(* IEC 61131-3 sources: 2026_Projet_YGO_ExcavatriceDragage/TOOLS/TEST_AUTO_CI/RESULTS/H_TREUILS_BENNE/tests (part 3) *)

(* ---- test_fb_winch.st ---- *)
(* =======================================================================
   🧪 test_fb_winch.st — FB_Winch (TC-P10-011, 017, 019, 042.1, 052.1, T216-AC4)
   ───────────────────────────────────────────────────────────────
   Fiche : DOC/AF/AF_Partie-10_Fonction_Winch/FB_Winch_v1.0.md
   Conventions : 1 appel fb() = 1 scan ; ADVANCE_TIME(10000000) entre les
   scans pour les fronts R_TRIG ; hex décrit en décimal (bit 0 = 1, bit 15 = 32768).
   Table valide : seuils croissants [10,30,50,70,90], P2..P5 au moins 1 contacteur TRUE.
   Interface structs : DriveRequest / Sensors / Config passés en variables
   (le harnais STruCpp ne supporte pas les littéraux de struct en appel FB).
   ======================================================================= *)

SETUP
VAR
    FB_W : FB_Winch;
    Table : ST_SpeedStepTable;
    DriveReq : ST_fbWinch_DriveRequest;
    Sens : ST_fbWinch_Sensors;
    Cfg : ST_fbWinch_Cfg;
END_VAR
END_SETUP

(* ── Table valide commune ── *)

TEST 'TC-P03-001 Dynamique Enable : neutralisation initiale, transition Ready au repos, puis coupure'
    Table.StepThreshold_Pct[1] := 10.0;
    Table.StepThreshold_Pct[2] := 30.0;
    Table.StepThreshold_Pct[3] := 50.0;
    Table.StepThreshold_Pct[4] := 70.0;
    Table.StepThreshold_Pct[5] := 90.0;
    Table.P2R1 := TRUE;
    Table.P3R1 := TRUE;
    Table.P4R1 := TRUE;
    Table.P5R1 := TRUE;
    Cfg.SpeedStepTable := Table;
    Sens.Homed := TRUE;
    Sens.ContactorsAllOff := TRUE;
    Sens.SpeedGuardReady := TRUE;

    (* Scan 0 : Enable=FALSE -> Neutralisation initiale *)
    DriveReq.RunRequest := FALSE;
    DriveReq.ReqAscent := FALSE; DriveReq.ReqDescend := FALSE;
    DriveReq.SpeedTgt_Pct := 0.0;
    FB_W(Enable := FALSE, Reset := FALSE, PowerContactorEngaged := TRUE,
         DriveRequest := DriveReq, Sensors := Sens, Config := Cfg);
    ASSERT_FALSE(FB_W.Ready, 'Enable=FALSE -> Ready=FALSE (neutralise)');

    ADVANCE_TIME(10000000);

    (* Scan 1 : Enable=TRUE -> Premier scan d initialisation *)
    FB_W(Enable := TRUE, Reset := FALSE, PowerContactorEngaged := TRUE,
         DriveRequest := DriveReq, Sensors := Sens, Config := Cfg);

    ADVANCE_TIME(10000000);

    (* Scan 2 : Regime nominal etabli -> Ready=TRUE *)
    FB_W(Enable := TRUE, Reset := FALSE, PowerContactorEngaged := TRUE,
         DriveRequest := DriveReq, Sensors := Sens, Config := Cfg);
    ASSERT_TRUE(FB_W.Ready, 'Enable=TRUE etabli -> Ready=TRUE (nominal)');

    ADVANCE_TIME(10000000);

    (* Scan 3 : Enable=FALSE -> Coupure nette et re-neutralisation *)
    FB_W(Enable := FALSE, Reset := FALSE, PowerContactorEngaged := TRUE,
         DriveRequest := DriveReq, Sensors := Sens, Config := Cfg);
    ASSERT_FALSE(FB_W.Ready, 'Enable=FALSE -> Ready retombe a FALSE');
END_TEST

TEST 'TC-P10-011 Inversion Fwd<->Rev : neutre->sens immediat, inversion exige delai + rampe a 0'
    Table.StepThreshold_Pct[1] := 10.0;
    Table.StepThreshold_Pct[2] := 30.0;
    Table.StepThreshold_Pct[3] := 50.0;
    Table.StepThreshold_Pct[4] := 70.0;
    Table.StepThreshold_Pct[5] := 90.0;
    Table.P2R1 := TRUE;
    Table.P3R1 := TRUE;
    Table.P4R1 := TRUE;
    Table.P5R1 := TRUE;
    Cfg.SpeedStepTable := Table;
    Sens.Homed := TRUE;
    Sens.ContactorsAllOff := TRUE;
    Sens.SpeedGuardReady := TRUE;

    (* Scan 1 : regime nominal *)
    DriveReq.RunRequest := FALSE;
    DriveReq.ReqAscent := FALSE; DriveReq.ReqDescend := FALSE;
    DriveReq.SpeedTgt_Pct := 0.0;
    FB_W(Enable := TRUE, Reset := FALSE, PowerContactorEngaged := TRUE,
         DriveRequest := DriveReq, Sensors := Sens, Config := Cfg);
    ADVANCE_TIME(10000000);
    FB_W(Enable := TRUE, Reset := FALSE, PowerContactorEngaged := TRUE,
         DriveRequest := DriveReq, Sensors := Sens, Config := Cfg);
    ASSERT_TRUE(FB_W.Ready, 'Treuil pret');

    (* Scan 2 : neutre -> montee = IMMEDIAT (pas de DirectionChangePending) *)
    ADVANCE_TIME(10000000);
    DriveReq.RunRequest := TRUE;
    DriveReq.ReqAscent := TRUE; DriveReq.ReqDescend := FALSE;
    DriveReq.SpeedTgt_Pct := 20.0;
    FB_W(Enable := TRUE, Reset := FALSE, PowerContactorEngaged := TRUE,
         DriveRequest := DriveReq, Sensors := Sens, Config := Cfg);
    ASSERT_EQ(FB_W.CommandedDirection, 1, 'Neutre->montee : CommandedDirection=1 immediat');
    ASSERT_FALSE(FB_W.DirectionChangePending, 'Neutre->montee : pas de pending');
    ASSERT_TRUE(FB_W.RelayFwd, 'Montee -> RelayFwd');

    (* Scan 3 : arret reel via neutre (StartStop=FALSE, Direction=0) -> StepNumber=0,
       CommandedDirection=0 (relais/diagnostic neutres) ; le dernier sens non nul est
       memorise en interne (LastDirection) pour l'interlock de reprise opposee *)
    ADVANCE_TIME(10000000);
    DriveReq.RunRequest := FALSE;
    DriveReq.ReqAscent := FALSE; DriveReq.ReqDescend := FALSE;
    DriveReq.SpeedTgt_Pct := 0.0;
    FB_W(Enable := TRUE, Reset := FALSE, PowerContactorEngaged := TRUE,
         DriveRequest := DriveReq, Sensors := Sens, Config := Cfg);
    ASSERT_EQ(FB_W.StepNumber, 0, 'Arret -> StepNumber=0');
    ASSERT_EQ(FB_W.CommandedDirection, 0, 'Arret via neutre : CommandedDirection=0 (relais/diagnostic neutres)');

    (* Scan 4 : inversion montee->descente apres neutre (StepNumber=0) -> pending + rampe a 0 *)
    ADVANCE_TIME(10000000);
    DriveReq.RunRequest := TRUE;
    DriveReq.ReqAscent := FALSE; DriveReq.ReqDescend := TRUE;
    DriveReq.SpeedTgt_Pct := 20.0;
    FB_W(Enable := TRUE, Reset := FALSE, PowerContactorEngaged := TRUE,
         DriveRequest := DriveReq, Sensors := Sens, Config := Cfg);
    ASSERT_TRUE(FB_W.DirectionChangePending, 'Inversion apres neutre -> DirectionChangePending=TRUE');
    ASSERT_EQ(FB_W.StepNumber, 0, 'Inversion : rampe forcee a 0 pendant attente');

    (* Scan 5 : apres DirectionInterlockDelayDescent=400ms -> CommandedDirection=-1 *)
    ADVANCE_TIME(400000000);
    FB_W(Enable := TRUE, Reset := FALSE, PowerContactorEngaged := TRUE,
         DriveRequest := DriveReq, Sensors := Sens, Config := Cfg);
    ASSERT_EQ(FB_W.CommandedDirection, -1, 'Apres 400ms -> CommandedDirection=-1');
    ASSERT_FALSE(FB_W.DirectionChangePending, 'Apres delai -> pending leve');
END_TEST

TEST 'TC-P10-011b Inversion via neutre : montee reelle -> relache neutre -> reprise descente -> temps mort + zero relais'
    Table.StepThreshold_Pct[1] := 10.0;
    Table.StepThreshold_Pct[2] := 30.0;
    Table.StepThreshold_Pct[3] := 50.0;
    Table.StepThreshold_Pct[4] := 70.0;
    Table.StepThreshold_Pct[5] := 90.0;
    Table.P2R1 := TRUE;
    Table.P3R1 := TRUE;
    Table.P4R1 := TRUE;
    Table.P5R1 := TRUE;
    Cfg.SpeedStepTable := Table;
    Sens.Homed := TRUE;
    Sens.ContactorsAllOff := TRUE;
    Sens.SpeedGuardReady := TRUE;

    (* Scan 1 : regime nominal *)
    DriveReq.RunRequest := FALSE;
    DriveReq.ReqAscent := FALSE; DriveReq.ReqDescend := FALSE;
    DriveReq.SpeedTgt_Pct := 0.0;
    FB_W(Enable := TRUE, Reset := FALSE, PowerContactorEngaged := TRUE,
         DriveRequest := DriveReq, Sensors := Sens, Config := Cfg);
    ADVANCE_TIME(10000000);
    FB_W(Enable := TRUE, Reset := FALSE, PowerContactorEngaged := TRUE,
         DriveRequest := DriveReq, Sensors := Sens, Config := Cfg);
    ASSERT_TRUE(FB_W.Ready, 'Treuil pret');

    (* Scan 2 : montee reelle etablie *)
    ADVANCE_TIME(10000000);
    DriveReq.RunRequest := TRUE;
    DriveReq.ReqAscent := TRUE; DriveReq.ReqDescend := FALSE;
    DriveReq.SpeedTgt_Pct := 90.0;
    FB_W(Enable := TRUE, Reset := FALSE, PowerContactorEngaged := TRUE,
         DriveRequest := DriveReq, Sensors := Sens, Config := Cfg);
    ASSERT_EQ(FB_W.CommandedDirection, 1, 'Montee reelle : CommandedDirection=1');
    ASSERT_TRUE(FB_W.RelayFwd, 'Montee reelle -> RelayFwd');

    (* Scan 3 : relachement neutre (Direction=0) -> StepNumber=0, CommandedDirection=0,
       relais coupes immediatement *)
    ADVANCE_TIME(10000000);
    DriveReq.RunRequest := FALSE;
    DriveReq.ReqAscent := FALSE; DriveReq.ReqDescend := FALSE;
    DriveReq.SpeedTgt_Pct := 0.0;
    FB_W(Enable := TRUE, Reset := FALSE, PowerContactorEngaged := TRUE,
         DriveRequest := DriveReq, Sensors := Sens, Config := Cfg);
    ASSERT_EQ(FB_W.StepNumber, 0, 'Neutre -> StepNumber=0');
    ASSERT_EQ(FB_W.CommandedDirection, 0, 'Neutre -> CommandedDirection=0 (relais/diagnostic neutres)');
    ASSERT_FALSE(FB_W.RelayFwd, 'Neutre -> RelayFwd coupe immediatement');
    ASSERT_FALSE(FB_W.RelayRev, 'Neutre -> RelayRev reste FALSE');

    (* Scan 4 : reprise descente (Direction=-1) -> pending + zero relais jusqu au delai *)
    ADVANCE_TIME(10000000);
    DriveReq.RunRequest := TRUE;
    DriveReq.ReqAscent := FALSE; DriveReq.ReqDescend := TRUE;
    DriveReq.SpeedTgt_Pct := 20.0;
    FB_W(Enable := TRUE, Reset := FALSE, PowerContactorEngaged := TRUE,
         DriveRequest := DriveReq, Sensors := Sens, Config := Cfg);
    ASSERT_TRUE(FB_W.DirectionChangePending, 'Reprise opposee apres neutre -> pending');
    ASSERT_EQ(FB_W.StepNumber, 0, 'Reprise opposee -> StepNumber=0 (rampe a 0)');
    ASSERT_FALSE(FB_W.RelayRev, 'Reprise opposee -> RelayRev retenu jusqu au delai');

    (* Scan 5 : apres DirectionInterlockDelayDescent=400ms -> CommandedDirection=-1, RelayRev *)
    ADVANCE_TIME(400000000);
    FB_W(Enable := TRUE, Reset := FALSE, PowerContactorEngaged := TRUE,
         DriveRequest := DriveReq, Sensors := Sens, Config := Cfg);
    ASSERT_EQ(FB_W.CommandedDirection, -1, 'Apres delai -> CommandedDirection=-1');
    ASSERT_FALSE(FB_W.DirectionChangePending, 'Apres delai -> pending leve');
    ASSERT_TRUE(FB_W.RelayRev, 'Apres delai -> RelayRev commande');
END_TEST

TEST 'TC-P10-011c Reprise du MEME sens apres neutre : depart immediat (pas de pending)'
    Table.StepThreshold_Pct[1] := 10.0;
    Table.StepThreshold_Pct[2] := 30.0;
    Table.StepThreshold_Pct[3] := 50.0;
    Table.StepThreshold_Pct[4] := 70.0;
    Table.StepThreshold_Pct[5] := 90.0;
    Table.P2R1 := TRUE;
    Table.P3R1 := TRUE;
    Table.P4R1 := TRUE;
    Table.P5R1 := TRUE;
    Cfg.SpeedStepTable := Table;
    Sens.Homed := TRUE;
    Sens.ContactorsAllOff := TRUE;
    Sens.SpeedGuardReady := TRUE;

    (* Scan 1 : regime nominal *)
    DriveReq.RunRequest := FALSE;
    DriveReq.ReqAscent := FALSE; DriveReq.ReqDescend := FALSE;
    DriveReq.SpeedTgt_Pct := 0.0;
    FB_W(Enable := TRUE, Reset := FALSE, PowerContactorEngaged := TRUE,
         DriveRequest := DriveReq, Sensors := Sens, Config := Cfg);
    ADVANCE_TIME(10000000);
    FB_W(Enable := TRUE, Reset := FALSE, PowerContactorEngaged := TRUE,
         DriveRequest := DriveReq, Sensors := Sens, Config := Cfg);
    ASSERT_TRUE(FB_W.Ready, 'Treuil pret');

    (* Scan 2 : montee reelle etablie *)
    ADVANCE_TIME(10000000);
    DriveReq.RunRequest := TRUE;
    DriveReq.ReqAscent := TRUE; DriveReq.ReqDescend := FALSE;
    DriveReq.SpeedTgt_Pct := 20.0;
    FB_W(Enable := TRUE, Reset := FALSE, PowerContactorEngaged := TRUE,
         DriveRequest := DriveReq, Sensors := Sens, Config := Cfg);
    ASSERT_EQ(FB_W.CommandedDirection, 1, 'Montee reelle : CommandedDirection=1');
    ASSERT_TRUE(FB_W.RelayFwd, 'Montee reelle -> RelayFwd');

    (* Scan 3 : relachement neutre -> CommandedDirection=0 *)
    ADVANCE_TIME(10000000);
    DriveReq.RunRequest := FALSE;
    DriveReq.ReqAscent := FALSE; DriveReq.ReqDescend := FALSE;
    DriveReq.SpeedTgt_Pct := 0.0;
    FB_W(Enable := TRUE, Reset := FALSE, PowerContactorEngaged := TRUE,
         DriveRequest := DriveReq, Sensors := Sens, Config := Cfg);
    ASSERT_EQ(FB_W.CommandedDirection, 0, 'Neutre -> CommandedDirection=0');

    (* Scan 4 : reprise du MEME sens (montee) -> depart immediat, pas de pending *)
    ADVANCE_TIME(10000000);
    DriveReq.RunRequest := TRUE;
    DriveReq.ReqAscent := TRUE; DriveReq.ReqDescend := FALSE;
    DriveReq.SpeedTgt_Pct := 20.0;
    FB_W(Enable := TRUE, Reset := FALSE, PowerContactorEngaged := TRUE,
         DriveRequest := DriveReq, Sensors := Sens, Config := Cfg);
    ASSERT_EQ(FB_W.CommandedDirection, 1, 'Reprise meme sens -> CommandedDirection=1 immediat');
    ASSERT_FALSE(FB_W.DirectionChangePending, 'Reprise meme sens -> pas de pending');
    ASSERT_TRUE(FB_W.RelayFwd, 'Reprise meme sens -> RelayFwd immediat');
END_TEST

TEST 'TC-P10-017 Config palier invalide : palier 0, sorties sures'
    (* Table invalide : seuils non croissants (tous a 0) *)
    Table.StepThreshold_Pct[1] := 0.0;
    Table.StepThreshold_Pct[2] := 0.0;
    Table.StepThreshold_Pct[3] := 0.0;
    Table.StepThreshold_Pct[4] := 0.0;
    Table.StepThreshold_Pct[5] := 0.0;
    Cfg.SpeedStepTable := Table;
    Sens.Homed := TRUE;
    Sens.ContactorsAllOff := TRUE;
    Sens.SpeedGuardReady := TRUE;

    (* Scan 1 : Enable=TRUE, config invalide -> ConfigError latche *)
    DriveReq.RunRequest := TRUE;
    DriveReq.ReqAscent := TRUE; DriveReq.ReqDescend := FALSE;
    DriveReq.SpeedTgt_Pct := 50.0;
    FB_W(Enable := TRUE, Reset := FALSE, PowerContactorEngaged := TRUE,
         DriveRequest := DriveReq, Sensors := Sens, Config := Cfg);
    ADVANCE_TIME(10000000);
    FB_W(Enable := TRUE, Reset := FALSE, PowerContactorEngaged := TRUE,
         DriveRequest := DriveReq, Sensors := Sens, Config := Cfg);
    ASSERT_TRUE(FB_W.Fault.Error, 'Config invalide -> Error');
    ASSERT_EQ(FB_W.StepNumber, 0, 'Config invalide -> palier 0');
    ASSERT_FALSE(FB_W.RelayFwd, 'Config invalide -> RelayFwd=FALSE (sortie sure)');
    ASSERT_FALSE(FB_W.RelayRev, 'Config invalide -> RelayRev=FALSE');
    ASSERT_FALSE(FB_W.Contactor1, 'Config invalide -> Contactor1=FALSE');
END_TEST

(* TC-P10-018 (StuckClosed) deplace/adapte dans test_fb_safety_winch.st (T181-02/03 AC5) :
   FB_Winch ne produit plus la detection contacteur colle — proprietaire unique FB_Safety_Winch. *)

TEST 'TC-P10-019 Ordre MainTask : Safety -> WinchControl -> PRG_06_Outputs'
    (* (essai site — stub) : l ordre d execution MainTask (Safety -> WinchControl -> PRG_06)
       est une propriete de la tache CODESYS, non automatisable en boite noire FB. On verifie
       ici la brique amont : FB_Winch produit bien sa demande sortie (RelayFwd) qui sera
       consommee par la barriere finale PRG_06. *)
    Table.StepThreshold_Pct[1] := 10.0;
    Table.StepThreshold_Pct[2] := 30.0;
    Table.StepThreshold_Pct[3] := 50.0;
    Table.StepThreshold_Pct[4] := 70.0;
    Table.StepThreshold_Pct[5] := 90.0;
    Table.P2R1 := TRUE;
    Table.P3R1 := TRUE;
    Table.P4R1 := TRUE;
    Table.P5R1 := TRUE;
    Cfg.SpeedStepTable := Table;
    Sens.Homed := TRUE;
    Sens.ContactorsAllOff := TRUE;
    Sens.SpeedGuardReady := TRUE;

    DriveReq.RunRequest := FALSE;
    DriveReq.ReqAscent := FALSE; DriveReq.ReqDescend := FALSE;
    DriveReq.SpeedTgt_Pct := 0.0;
    FB_W(Enable := TRUE, Reset := FALSE, PowerContactorEngaged := TRUE,
         DriveRequest := DriveReq, Sensors := Sens, Config := Cfg);
    ADVANCE_TIME(10000000);
    DriveReq.RunRequest := TRUE;
    DriveReq.ReqAscent := TRUE; DriveReq.ReqDescend := FALSE;
    DriveReq.SpeedTgt_Pct := 20.0;
    FB_W(Enable := TRUE, Reset := FALSE, PowerContactorEngaged := TRUE,
         DriveRequest := DriveReq, Sensors := Sens, Config := Cfg);
    ASSERT_TRUE(FB_W.RelayFwd, 'Demande montee produite (consommee par PRG_06)');
    ASSERT_TRUE(FB_W.Contactor1, 'Palier 1 demande');
END_TEST

TEST 'TC-P10-042.1 Plafonds dynamiques palier : descente max 3, montee max 5, approche capteur haut=1'
    Table.StepThreshold_Pct[1] := 10.0;
    Table.StepThreshold_Pct[2] := 30.0;
    Table.StepThreshold_Pct[3] := 50.0;
    Table.StepThreshold_Pct[4] := 70.0;
    Table.StepThreshold_Pct[5] := 90.0;
    Table.P2R1 := TRUE;
    Table.P3R1 := TRUE;
    Table.P4R1 := TRUE;
    Table.P5R1 := TRUE;
    Cfg.SpeedStepTable := Table;
    Sens.Homed := TRUE;
    Sens.ContactorsAllOff := TRUE;
    Sens.SpeedGuardReady := TRUE;
    DriveReq.HomingApproachActive := FALSE;
    Sens.CablePosM := 0.0;
    Cfg.SlowdownDistance_M := 1.0;

    (* Scan 1 : regime nominal *)
    DriveReq.RunRequest := FALSE;
    DriveReq.ReqAscent := FALSE; DriveReq.ReqDescend := FALSE;
    DriveReq.SpeedTgt_Pct := 0.0;
    FB_W(Enable := TRUE, Reset := FALSE, PowerContactorEngaged := TRUE,
         DriveRequest := DriveReq, Sensors := Sens, Config := Cfg);
    ADVANCE_TIME(10000000);
    FB_W(Enable := TRUE, Reset := FALSE, PowerContactorEngaged := TRUE,
         DriveRequest := DriveReq, Sensors := Sens, Config := Cfg);

    (* Descente : SpeedTgt_Pct=90 -> RequestedStep cape a CfgMaxStepDescente=3 *)
    ADVANCE_TIME(10000000);
    DriveReq.RunRequest := TRUE;
    DriveReq.ReqAscent := FALSE; DriveReq.ReqDescend := TRUE;
    DriveReq.SpeedTgt_Pct := 90.0;
    FB_W(Enable := TRUE, Reset := FALSE, PowerContactorEngaged := TRUE,
         DriveRequest := DriveReq, Sensors := Sens, Config := Cfg);
    ASSERT_EQ(FB_W.RequestedStep, 3, 'Descente : palier cape a 3 (CfgMaxStepDescente)');

    (* Reset + montee : SpeedTgt_Pct=90 -> RequestedStep=5 (MaxStepAscent) *)
    ADVANCE_TIME(10000000);
    DriveReq.RunRequest := FALSE;
    DriveReq.ReqAscent := FALSE; DriveReq.ReqDescend := FALSE;
    DriveReq.SpeedTgt_Pct := 0.0;
    FB_W(Enable := TRUE, Reset := TRUE, PowerContactorEngaged := TRUE,
         DriveRequest := DriveReq, Sensors := Sens, Config := Cfg);
    ADVANCE_TIME(10000000);
    DriveReq.RunRequest := TRUE;
    DriveReq.ReqAscent := TRUE; DriveReq.ReqDescend := FALSE;
    DriveReq.SpeedTgt_Pct := 90.0;
    FB_W(Enable := TRUE, Reset := FALSE, PowerContactorEngaged := TRUE,
         DriveRequest := DriveReq, Sensors := Sens, Config := Cfg);
    ASSERT_EQ(FB_W.RequestedStep, 5, 'Montee : palier 5 (MaxStepAscent)');

    (* Approche capteur haut : HomingApproachActive=TRUE -> palier 1 *)
    ADVANCE_TIME(10000000);
    DriveReq.RunRequest := FALSE;
    DriveReq.ReqAscent := FALSE; DriveReq.ReqDescend := FALSE;
    DriveReq.SpeedTgt_Pct := 0.0;
    FB_W(Enable := TRUE, Reset := TRUE, PowerContactorEngaged := TRUE,
         DriveRequest := DriveReq, Sensors := Sens, Config := Cfg);
    ADVANCE_TIME(10000000);
    DriveReq.RunRequest := TRUE;
    DriveReq.ReqAscent := TRUE; DriveReq.ReqDescend := FALSE;
    DriveReq.SpeedTgt_Pct := 90.0;
    DriveReq.HomingApproachActive := TRUE;
    FB_W(Enable := TRUE, Reset := FALSE, PowerContactorEngaged := TRUE,
         DriveRequest := DriveReq, Sensors := Sens, Config := Cfg);
    ASSERT_EQ(FB_W.RequestedStep, 1, 'Approche capteur haut : palier 1');

    (* Zone ralentissement haut : CablePosM >= TopLimitM - CfgSlowdownDistanceM -> palier 1 *)
    ADVANCE_TIME(10000000);
    DriveReq.RunRequest := FALSE;
    DriveReq.ReqAscent := FALSE; DriveReq.ReqDescend := FALSE;
    DriveReq.SpeedTgt_Pct := 0.0;
    DriveReq.HomingApproachActive := FALSE;
    FB_W(Enable := TRUE, Reset := TRUE, PowerContactorEngaged := TRUE,
         DriveRequest := DriveReq, Sensors := Sens, Config := Cfg);
    ADVANCE_TIME(10000000);
    DriveReq.RunRequest := TRUE;
    DriveReq.ReqAscent := TRUE; DriveReq.ReqDescend := FALSE;
    DriveReq.SpeedTgt_Pct := 90.0;
    DriveReq.TopLimitM := 8.5;
    Sens.CablePosM := 8.0;
    Cfg.SlowdownDistance_M := 1.0;
    FB_W(Enable := TRUE, Reset := FALSE, PowerContactorEngaged := TRUE,
         DriveRequest := DriveReq, Sensors := Sens, Config := Cfg);
    ASSERT_TRUE(FB_W.InTopSlowdownZone, 'Zone ralentissement haut active');
    ASSERT_EQ(FB_W.RequestedStep, 1, 'Zone ralentissement haut : palier 1');
END_TEST

TEST 'TC-P10-052.1 Garde-fou vitesse : vitesse non-stable -> palier 1 (activation par defaut)'
    (* (activation par defaut : T177) — SpeedGuardEnable est TRUE par defaut dans le code.
       On ne le force pas : le test verifie que le garde-fou est actif sans activation manuelle. *)
    Table.StepThreshold_Pct[1] := 10.0;
    Table.StepThreshold_Pct[2] := 30.0;
    Table.StepThreshold_Pct[3] := 50.0;
    Table.StepThreshold_Pct[4] := 70.0;
    Table.StepThreshold_Pct[5] := 90.0;
    Table.P2R1 := TRUE;
    Table.P3R1 := TRUE;
    Table.P4R1 := TRUE;
    Table.P5R1 := TRUE;
    Cfg.SpeedStepTable := Table;
    Sens.Homed := TRUE;
    Sens.ContactorsAllOff := TRUE;
    Sens.SpeedGuardReady := TRUE;
    DriveReq.HomingApproachActive := FALSE;
    Sens.CablePosM := 0.0;
    Cfg.SlowdownDistance_M := 1.0;

    (* Scan 1 : regime nominal *)
    DriveReq.RunRequest := FALSE;
    DriveReq.ReqAscent := FALSE; DriveReq.ReqDescend := FALSE;
    DriveReq.SpeedTgt_Pct := 0.0;
    FB_W(Enable := TRUE, Reset := FALSE, PowerContactorEngaged := TRUE,
         DriveRequest := DriveReq, Sensors := Sens, Config := Cfg);
    ADVANCE_TIME(10000000);
    FB_W(Enable := TRUE, Reset := FALSE, PowerContactorEngaged := TRUE,
         DriveRequest := DriveReq, Sensors := Sens, Config := Cfg);

    (* Scan 2 : SpeedGuardEnable=TRUE (defaut), SpeedGuardReady=FALSE (vitesse non stable) -> palier 1 *)
    ADVANCE_TIME(10000000);
    DriveReq.RunRequest := TRUE;
    DriveReq.ReqAscent := TRUE; DriveReq.ReqDescend := FALSE;
    DriveReq.SpeedTgt_Pct := 90.0;
    Sens.SpeedGuardReady := FALSE;
    FB_W(Enable := TRUE, Reset := FALSE, PowerContactorEngaged := TRUE,
         DriveRequest := DriveReq, Sensors := Sens, Config := Cfg);
    ASSERT_EQ(FB_W.RequestedStep, 1, 'Vitesse non stable -> palier 1 (garde-fou)');
    ASSERT_EQ(FB_W.StepNumber, 1, 'Vitesse non stable -> StepNumber=1');
END_TEST

(* ───────────────────────────────────────────────────────────────
   T216-AC4 : le plancher MinStepDown ne relance JAMAIS une descente
   lorsque le permis effectif de descente est FALSE (EffectiveSafeStop).
   REX : limite basse atteinte -> DescendPermit=FALSE -> la descente
   continuait au palier 1 (relance physique). Correction : gate du
   plancher par NOT EffectiveSafeStop (ligne 242 FB_Winch.st).
   ─────────────────────────────────────────────────────────────── *)

TEST 'T216-AC4-1 Regression : DescendPermit=FALSE + MinStepDown=1 -> StepNumber=0 et sorties=0'
    Table.StepThreshold_Pct[1] := 10.0;
    Table.StepThreshold_Pct[2] := 30.0;
    Table.StepThreshold_Pct[3] := 50.0;
    Table.StepThreshold_Pct[4] := 70.0;
    Table.StepThreshold_Pct[5] := 90.0;
    Table.P2R1 := TRUE;
    Table.P3R1 := TRUE;
    Table.P4R1 := TRUE;
    Table.P5R1 := TRUE;
    Cfg.SpeedStepTable := Table;
    Sens.Homed := TRUE;
    Sens.ContactorsAllOff := TRUE;
    Sens.SpeedGuardReady := TRUE;
    DriveReq.HomingApproachActive := FALSE;
    Sens.CablePosM := 0.0;
    Cfg.SlowdownDistance_M := 1.0;

    // Scan 1 : regime nominal neutre (arme l interlock direction), permis deja FALSE
    DriveReq.RunRequest := FALSE;
    DriveReq.ReqAscent := FALSE; DriveReq.ReqDescend := FALSE;
    DriveReq.SpeedStepReq := 0;
    DriveReq.MinStepDown := 1;
    DriveReq.MaxStepDown := 3;
    FB_W(Enable := TRUE, Reset := FALSE, PowerContactorEngaged := TRUE,
         DriveRequest := DriveReq, Sensors := Sens, Config := Cfg,
         SafeStop := FALSE, DescendPermit := FALSE, AscentPermit := TRUE);
    ADVANCE_TIME(10000000);
    FB_W(Enable := TRUE, Reset := FALSE, PowerContactorEngaged := TRUE,
         DriveRequest := DriveReq, Sensors := Sens, Config := Cfg,
         SafeStop := FALSE, DescendPermit := FALSE, AscentPermit := TRUE);

    // Scan 2 : operateur demande la descente (StartStop=TRUE, Dir=-1, SpeedStepReq=1)
    // MAIS DescendPermit=FALSE -> EffectiveSafeStop=TRUE doit garder RequestedStep=0.
    // Le plancher MinStepDown=1 ne doit PAS relever RequestedStep a >=1.
    ADVANCE_TIME(10000000);
    DriveReq.RunRequest := TRUE;
    DriveReq.ReqAscent := FALSE; DriveReq.ReqDescend := TRUE;
    DriveReq.SpeedStepReq := 1;
    FB_W(Enable := TRUE, Reset := FALSE, PowerContactorEngaged := TRUE,
         DriveRequest := DriveReq, Sensors := Sens, Config := Cfg,
         SafeStop := FALSE, DescendPermit := FALSE, AscentPermit := TRUE);
    ASSERT_EQ(FB_W.StepNumber, 0, 'Permis FALSE + MinStepDown : StepNumber=0 (descente interdite)');
    ASSERT_FALSE(FB_W.RelayFwd, 'Permis FALSE -> RelayFwd=FALSE');
    ASSERT_FALSE(FB_W.RelayRev, 'Permis FALSE -> RelayRev=FALSE (aucune relance descente)');
    ASSERT_FALSE(FB_W.Contactor1, 'Permis FALSE -> Contactor1=FALSE (sorties DQ descente = 0)');

    // Scan 3..4 : la demande est maintenue -> aucune relance palier apres cadence
    ADVANCE_TIME(10000000);
    FB_W(Enable := TRUE, Reset := FALSE, PowerContactorEngaged := TRUE,
         DriveRequest := DriveReq, Sensors := Sens, Config := Cfg,
         SafeStop := FALSE, DescendPermit := FALSE, AscentPermit := TRUE);
    ADVANCE_TIME(500000000);
    FB_W(Enable := TRUE, Reset := FALSE, PowerContactorEngaged := TRUE,
         DriveRequest := DriveReq, Sensors := Sens, Config := Cfg,
         SafeStop := FALSE, DescendPermit := FALSE, AscentPermit := TRUE);
    ASSERT_EQ(FB_W.StepNumber, 0, 'Permis FALSE : StepNumber reste 0 apres cadence (aucune relance)');
    ASSERT_FALSE(FB_W.RelayRev, 'Permis FALSE : RelayRev reste FALSE apres cadence');
END_TEST

TEST 'T216-AC4-2 Non-regression plongee Kobold : DescendPermit=TRUE + MinStepDown=3 -> plancher applique'
    Table.StepThreshold_Pct[1] := 10.0;
    Table.StepThreshold_Pct[2] := 30.0;
    Table.StepThreshold_Pct[3] := 50.0;
    Table.StepThreshold_Pct[4] := 70.0;
    Table.StepThreshold_Pct[5] := 90.0;
    Table.P2R1 := TRUE;
    Table.P3R1 := TRUE;
    Table.P4R1 := TRUE;
    Table.P5R1 := TRUE;
    Cfg.SpeedStepTable := Table;
    Sens.Homed := TRUE;
    Sens.ContactorsAllOff := TRUE;
    Sens.SpeedGuardReady := TRUE;
    DriveReq.HomingApproachActive := FALSE;
    Sens.CablePosM := 0.0;
    Cfg.SlowdownDistance_M := 1.0;

    // Scan 1 : regime nominal neutre
    DriveReq.RunRequest := FALSE;
    DriveReq.ReqAscent := FALSE; DriveReq.ReqDescend := FALSE;
    DriveReq.SpeedStepReq := 0;
    DriveReq.MinStepDown := 3;
    DriveReq.MaxStepDown := 3;
    FB_W(Enable := TRUE, Reset := FALSE, PowerContactorEngaged := TRUE,
         DriveRequest := DriveReq, Sensors := Sens, Config := Cfg,
         SafeStop := FALSE, DescendPermit := TRUE, AscentPermit := TRUE);
    ADVANCE_TIME(10000000);
    FB_W(Enable := TRUE, Reset := FALSE, PowerContactorEngaged := TRUE,
         DriveRequest := DriveReq, Sensors := Sens, Config := Cfg,
         SafeStop := FALSE, DescendPermit := TRUE, AscentPermit := TRUE);

    // Scan 2 : descente demandee, cible basse (SpeedStepReq=1) mais plancher MinStepDown=3
    // permis OK -> le plancher releve RequestedStep a 3 (clamp au plafond MaxStepDown=3)
    ADVANCE_TIME(10000000);
    DriveReq.RunRequest := TRUE;
    DriveReq.ReqAscent := FALSE; DriveReq.ReqDescend := TRUE;
    DriveReq.SpeedStepReq := 1;
    FB_W(Enable := TRUE, Reset := FALSE, PowerContactorEngaged := TRUE,
         DriveRequest := DriveReq, Sensors := Sens, Config := Cfg,
         SafeStop := FALSE, DescendPermit := TRUE, AscentPermit := TRUE);
    ASSERT_EQ(FB_W.RequestedStep, 3, 'Plancher MinStepDown=3 releve RequestedStep (permis OK)');
    ASSERT_TRUE(FB_W.StepNumber > 0, 'Plancher MinStepDown=3 -> StepNumber>0 (plongee maintenue)');
    ASSERT_TRUE(FB_W.RelayRev, 'Plancher MinStepDown=3 -> RelayRev commande (plongee Kobold)');

    // Scan 3..4 : cadence des 2 crans suivants (500ms/cran descente) -> StepNumber=3
    ADVANCE_TIME(500000000);
    FB_W(Enable := TRUE, Reset := FALSE, PowerContactorEngaged := TRUE,
         DriveRequest := DriveReq, Sensors := Sens, Config := Cfg,
         SafeStop := FALSE, DescendPermit := TRUE, AscentPermit := TRUE);
    ADVANCE_TIME(500000000);
    FB_W(Enable := TRUE, Reset := FALSE, PowerContactorEngaged := TRUE,
         DriveRequest := DriveReq, Sensors := Sens, Config := Cfg,
         SafeStop := FALSE, DescendPermit := TRUE, AscentPermit := TRUE);
    ASSERT_EQ(FB_W.StepNumber, 3, 'Cadence complet -> StepNumber=3 (plancher + plafond clamp)');
END_TEST

TEST 'T216-AC4-3 Perte du permis en mouvement : StepNumber retombe a 0 sans reprise de plancher'
    Table.StepThreshold_Pct[1] := 10.0;
    Table.StepThreshold_Pct[2] := 30.0;
    Table.StepThreshold_Pct[3] := 50.0;
    Table.StepThreshold_Pct[4] := 70.0;
    Table.StepThreshold_Pct[5] := 90.0;
    Table.P2R1 := TRUE;
    Table.P3R1 := TRUE;
    Table.P4R1 := TRUE;
    Table.P5R1 := TRUE;
    Cfg.SpeedStepTable := Table;
    Sens.Homed := TRUE;
    Sens.ContactorsAllOff := TRUE;
    Sens.SpeedGuardReady := TRUE;
    DriveReq.HomingApproachActive := FALSE;
    Sens.CablePosM := 0.0;
    Cfg.SlowdownDistance_M := 1.0;

    // Scan 1 : regime nominal neutre
    DriveReq.RunRequest := FALSE;
    DriveReq.ReqAscent := FALSE; DriveReq.ReqDescend := FALSE;
    DriveReq.SpeedStepReq := 0;
    DriveReq.MinStepDown := 1;
    DriveReq.MaxStepDown := 3;
    FB_W(Enable := TRUE, Reset := FALSE, PowerContactorEngaged := TRUE,
         DriveRequest := DriveReq, Sensors := Sens, Config := Cfg,
         SafeStop := FALSE, DescendPermit := TRUE, AscentPermit := TRUE);
    ADVANCE_TIME(10000000);
    FB_W(Enable := TRUE, Reset := FALSE, PowerContactorEngaged := TRUE,
         DriveRequest := DriveReq, Sensors := Sens, Config := Cfg,
         SafeStop := FALSE, DescendPermit := TRUE, AscentPermit := TRUE);

    // Scan 2-3 : descente etablie (permis OK) -> StepNumber=1, RelayRev commande
    ADVANCE_TIME(10000000);
    DriveReq.RunRequest := TRUE;
    DriveReq.ReqAscent := FALSE; DriveReq.ReqDescend := TRUE;
    DriveReq.SpeedStepReq := 1;
    FB_W(Enable := TRUE, Reset := FALSE, PowerContactorEngaged := TRUE,
         DriveRequest := DriveReq, Sensors := Sens, Config := Cfg,
         SafeStop := FALSE, DescendPermit := TRUE, AscentPermit := TRUE);
    ADVANCE_TIME(10000000);
    FB_W(Enable := TRUE, Reset := FALSE, PowerContactorEngaged := TRUE,
         DriveRequest := DriveReq, Sensors := Sens, Config := Cfg,
         SafeStop := FALSE, DescendPermit := TRUE, AscentPermit := TRUE);
    ASSERT_TRUE(FB_W.RelayRev, 'Pre-condition : descente etablie (permis OK)');

    // Scan 4..6 : le permis descente TOMBE (limite basse atteinte), l operateur maintient
    // la demande (StartStop=TRUE, Dir=-1, MinStepDown=1) -> StepNumber doit retomber a 0
    ADVANCE_TIME(10000000);
    FB_W(Enable := TRUE, Reset := FALSE, PowerContactorEngaged := TRUE,
         DriveRequest := DriveReq, Sensors := Sens, Config := Cfg,
         SafeStop := FALSE, DescendPermit := FALSE, AscentPermit := TRUE);
    ADVANCE_TIME(10000000);
    FB_W(Enable := TRUE, Reset := FALSE, PowerContactorEngaged := TRUE,
         DriveRequest := DriveReq, Sensors := Sens, Config := Cfg,
         SafeStop := FALSE, DescendPermit := FALSE, AscentPermit := TRUE);
    ADVANCE_TIME(10000000);
    FB_W(Enable := TRUE, Reset := FALSE, PowerContactorEngaged := TRUE,
         DriveRequest := DriveReq, Sensors := Sens, Config := Cfg,
         SafeStop := FALSE, DescendPermit := FALSE, AscentPermit := TRUE);
    ASSERT_EQ(FB_W.StepNumber, 0, 'Permis tombe en mouvement -> StepNumber retombe a 0');
    ASSERT_FALSE(FB_W.RelayRev, 'Permis tombe en mouvement -> RelayRev=FALSE (interruption descente)');

    // Scan 7-8 : maintien de la demande sans reprise -> aucune re-atterrissage palier
    ADVANCE_TIME(500000000);
    FB_W(Enable := TRUE, Reset := FALSE, PowerContactorEngaged := TRUE,
         DriveRequest := DriveReq, Sensors := Sens, Config := Cfg,
         SafeStop := FALSE, DescendPermit := FALSE, AscentPermit := TRUE);
    ADVANCE_TIME(500000000);
    FB_W(Enable := TRUE, Reset := FALSE, PowerContactorEngaged := TRUE,
         DriveRequest := DriveReq, Sensors := Sens, Config := Cfg,
         SafeStop := FALSE, DescendPermit := FALSE, AscentPermit := TRUE);
    ASSERT_EQ(FB_W.StepNumber, 0, 'Permis tombe : StepNumber reste 0 apres cadence (pas de reprise)');
    ASSERT_FALSE(FB_W.RelayRev, 'Permis tombe : RelayRev reste FALSE apres cadence');
END_TEST

(* ---- test_fb_winch_speed_learning.st ---- *)
(* =======================================================================
   🧪 test_fb_winch_speed_learning.st — FB_WinchSpeedLearning (T181-15)
   ───────────────────────────────────────────────────────────────
   Collecteur STRICTEMENT PASSIF des vitesses reelles par palier (RETAIN).
   Contrat : DOC/WFLOW/CONTRACTS/TASK_CONTRACT_T181-15_SPEED_LEARNING.yaml
   Conventions : 1 appel fb() = 1 scan ; Table est VAR_IN_OUT.
   ✅ Harnais copy-out (T181-21) : run_tests.py injecte le copy-out des
   VAR_IN_OUT apres chaque fb() (inject_var_in_out_copyout.py) — la variable
   de test Table reflete donc les ecritures du FB apres l'appel. On peut
   desormais asserter sur Table.Cell[...] (moyenne glissante + persistance
   RETAIN, TC-T181-15j).
   Strategie : pre-remplir la variable de test Table AVANT fb() pour les
   tests de frontiere/completude (a..i), et asserter sur Table.Cell[...]
   apres fb() pour prouver la moyenne glissante et la persistance RETAIN (j).
   Passivite (AC1/AC7) : verifiee par grep de l'interface FB (aucune sortie
   actionneur Relay* / Contactor* / Brake* / SpeedCmd ni Overspeed* / SpeedGuard* ).
   ======================================================================= *)

SETUP
VAR
    fb : FB_WinchSpeedLearning;
    Table : ST_fbWinchSpeedLearning_Table;
    Cfg : ST_fbWinchSpeedLearning_Cfg;
END_VAR
END_SETUP

(* ── Config commune : enveloppes par palier + MinSamples=3 ── *)

TEST 'TC-T181-15a LearnStart=FALSE : aucune collecte, table inchangee (AC3)'
    Cfg.MinSpeedMps[1] := 0.5; Cfg.MaxSpeedMps[1] := 2.0;
    Cfg.MinSpeedMps[2] := 1.0; Cfg.MaxSpeedMps[2] := 3.0;
    Cfg.MinSpeedMps[3] := 1.5; Cfg.MaxSpeedMps[3] := 4.0;
    Cfg.MinSpeedMps[4] := 2.0; Cfg.MaxSpeedMps[4] := 5.0;
    Cfg.MinSpeedMps[5] := 2.5; Cfg.MaxSpeedMps[5] := 6.0;
    Cfg.MinSamples := 3;

    (* Pre-remplissage : 1 cellule valide [1,1,1,1] *)
    Table.Cell[1][1][1][1].Valid := TRUE;
    Table.Cell[1][1][1][1].SpeedMps := 1.5;
    Table.Cell[1][1][1][1].SampleCount := 3;

    (* LearnStart=FALSE, toutes les autres conditions de collecte valides *)
    fb(Enable := TRUE, LearnStart := FALSE, WinchId := 1, Direction := 1,
       StepNumber := 1, MeasuredSpeedMps := 1.5, MeasuredSpeedValid := TRUE,
       LoadPresent := FALSE, StableForLearn := TRUE, Config := Cfg, Table := Table);

    ASSERT_FALSE(fb.Learning, 'LearnStart=FALSE : pas de collecte (Learning=FALSE)');
    ASSERT_FALSE(fb.LampLearn, 'LearnStart=FALSE : pas de voyant apprentissage');
    ASSERT_EQ(fb.CellsFilled, 1, 'LearnStart=FALSE : aucune nouvelle cellule (CellsFilled=1)');
END_TEST

TEST 'TC-T181-15b Conditions de collecte manquantes une a une : aucune ecriture (AC4)'
    Cfg.MinSpeedMps[1] := 0.5; Cfg.MaxSpeedMps[1] := 2.0;
    Cfg.MinSpeedMps[2] := 1.0; Cfg.MaxSpeedMps[2] := 3.0;
    Cfg.MinSpeedMps[3] := 1.5; Cfg.MaxSpeedMps[3] := 4.0;
    Cfg.MinSpeedMps[4] := 2.0; Cfg.MaxSpeedMps[4] := 5.0;
    Cfg.MinSpeedMps[5] := 2.5; Cfg.MaxSpeedMps[5] := 6.0;
    Cfg.MinSamples := 3;

    (* Mesure non valide : collecte bloquee -> aucune nouvelle cellule (CellsFilled reste 1) *)
    Table.Cell[1][1][1][1].Valid := TRUE;
    Table.Cell[1][1][1][1].SpeedMps := 1.5;
    Table.Cell[1][1][1][1].SampleCount := 3;
    fb(Enable := TRUE, LearnStart := TRUE, WinchId := 1, Direction := 1,
       StepNumber := 2, MeasuredSpeedMps := 1.5, MeasuredSpeedValid := FALSE,
       LoadPresent := FALSE, StableForLearn := TRUE, Config := Cfg, Table := Table);
    ASSERT_FALSE(fb.Learning, 'Mesure non valide : pas de collecte');
    ASSERT_EQ(fb.CellsFilled, 1, 'Mesure non valide : aucune nouvelle cellule');

    (* Conditions instables : collecte bloquee -> aucune nouvelle cellule *)
    Table.Cell[1][1][1][1].Valid := TRUE;
    Table.Cell[1][1][1][1].SpeedMps := 1.5;
    Table.Cell[1][1][1][1].SampleCount := 3;
    fb(Enable := TRUE, LearnStart := TRUE, WinchId := 1, Direction := 1,
       StepNumber := 3, MeasuredSpeedMps := 1.5, MeasuredSpeedValid := TRUE,
       LoadPresent := FALSE, StableForLearn := FALSE, Config := Cfg, Table := Table);
    ASSERT_FALSE(fb.Learning, 'Conditions instables : pas de collecte');
    ASSERT_EQ(fb.CellsFilled, 1, 'Conditions instables : aucune nouvelle cellule');

    (* Sens nul : collecte bloquee -> aucune nouvelle cellule *)
    Table.Cell[1][1][1][1].Valid := TRUE;
    Table.Cell[1][1][1][1].SpeedMps := 1.5;
    Table.Cell[1][1][1][1].SampleCount := 3;
    fb(Enable := TRUE, LearnStart := TRUE, WinchId := 1, Direction := 0,
       StepNumber := 4, MeasuredSpeedMps := 1.5, MeasuredSpeedValid := TRUE,
       LoadPresent := FALSE, StableForLearn := TRUE, Config := Cfg, Table := Table);
    ASSERT_FALSE(fb.Learning, 'Sens nul : pas de collecte');
    ASSERT_EQ(fb.CellsFilled, 1, 'Sens nul : aucune nouvelle cellule');

    (* Palier hors 1..5 : collecte bloquee -> aucune nouvelle cellule *)
    Table.Cell[1][1][1][1].Valid := TRUE;
    Table.Cell[1][1][1][1].SpeedMps := 1.5;
    Table.Cell[1][1][1][1].SampleCount := 3;
    fb(Enable := TRUE, LearnStart := TRUE, WinchId := 1, Direction := 1,
       StepNumber := 0, MeasuredSpeedMps := 1.5, MeasuredSpeedValid := TRUE,
       LoadPresent := FALSE, StableForLearn := TRUE, Config := Cfg, Table := Table);
    ASSERT_FALSE(fb.Learning, 'Palier hors 1..5 : pas de collecte');
    ASSERT_EQ(fb.CellsFilled, 1, 'Palier hors 1..5 : aucune nouvelle cellule');

    (* Axe hors 1..2 : collecte bloquee -> aucune nouvelle cellule *)
    Table.Cell[1][1][1][1].Valid := TRUE;
    Table.Cell[1][1][1][1].SpeedMps := 1.5;
    Table.Cell[1][1][1][1].SampleCount := 3;
    fb(Enable := TRUE, LearnStart := TRUE, WinchId := 0, Direction := 1,
       StepNumber := 1, MeasuredSpeedMps := 1.5, MeasuredSpeedValid := TRUE,
       LoadPresent := FALSE, StableForLearn := TRUE, Config := Cfg, Table := Table);
    ASSERT_FALSE(fb.Learning, 'Axe hors 1..2 : pas de collecte');
    ASSERT_EQ(fb.CellsFilled, 1, 'Axe hors 1..2 : aucune nouvelle cellule');
END_TEST

TEST 'TC-T181-15c Valid seulement a MinSamples : frontiere via CellsFilled (AC2/AC5)'
VAR
    i : INT;
    j : INT;
    k : INT;
    l : INT;
END_VAR
    Cfg.MinSpeedMps[1] := 0.5; Cfg.MaxSpeedMps[1] := 2.0;
    Cfg.MinSpeedMps[2] := 1.0; Cfg.MaxSpeedMps[2] := 3.0;
    Cfg.MinSpeedMps[3] := 1.5; Cfg.MaxSpeedMps[3] := 4.0;
    Cfg.MinSpeedMps[4] := 2.0; Cfg.MaxSpeedMps[4] := 5.0;
    Cfg.MinSpeedMps[5] := 2.5; Cfg.MaxSpeedMps[5] := 6.0;
    Cfg.MinSamples := 3;

    (* Part 1 : SampleCount=1 (MinSamples-2) -> apres 1 scan, encore < MinSamples -> non valide *)
    FOR i := 1 TO 2 DO
        FOR j := 1 TO 2 DO
            FOR k := 1 TO 2 DO
                FOR l := 1 TO 5 DO
                    Table.Cell[i][j][k][l].Valid := TRUE;
                END_FOR;
            END_FOR;
        END_FOR;
    END_FOR;
    Table.Cell[1][1][1][1].Valid := FALSE;
    Table.Cell[1][1][1][1].SampleCount := 1;
    Table.Cell[1][1][1][1].SpeedMps := 1.0;
    fb(Enable := TRUE, LearnStart := TRUE, WinchId := 1, Direction := 1,
       StepNumber := 1, MeasuredSpeedMps := 1.5, MeasuredSpeedValid := TRUE,
       LoadPresent := FALSE, StableForLearn := TRUE, Config := Cfg, Table := Table);
    ASSERT_EQ(fb.CellsFilled, 39, 'SampleCount 1->2 (<MinSamples) : cellule pas encore valide (39)');

    (* Part 2 : SampleCount=2 (MinSamples-1) -> apres 1 scan, MinSamples atteint -> valide *)
    FOR i := 1 TO 2 DO
        FOR j := 1 TO 2 DO
            FOR k := 1 TO 2 DO
                FOR l := 1 TO 5 DO
                    Table.Cell[i][j][k][l].Valid := TRUE;
                END_FOR;
            END_FOR;
        END_FOR;
    END_FOR;
    Table.Cell[1][1][1][1].Valid := FALSE;
    Table.Cell[1][1][1][1].SampleCount := 2;
    Table.Cell[1][1][1][1].SpeedMps := 1.0;
    fb(Enable := TRUE, LearnStart := TRUE, WinchId := 1, Direction := 1,
       StepNumber := 1, MeasuredSpeedMps := 1.5, MeasuredSpeedValid := TRUE,
       LoadPresent := FALSE, StableForLearn := TRUE, Config := Cfg, Table := Table);
    ASSERT_EQ(fb.CellsFilled, 40, 'SampleCount 2->3 (=MinSamples) : cellule validee (40)');
    ASSERT_TRUE(fb.TableComplete, 'MinSamples atteint sur la derniere cellule : TableComplete=TRUE');
END_TEST

TEST 'TC-T181-15d Hors enveloppe : cellule invalidee (Valid=FALSE, SampleCount=0, SpeedMps=0) (AC5)'
    Cfg.MinSpeedMps[1] := 0.5; Cfg.MaxSpeedMps[1] := 2.0;
    Cfg.MinSpeedMps[2] := 1.0; Cfg.MaxSpeedMps[2] := 3.0;
    Cfg.MinSpeedMps[3] := 1.5; Cfg.MaxSpeedMps[3] := 4.0;
    Cfg.MinSpeedMps[4] := 2.0; Cfg.MaxSpeedMps[4] := 5.0;
    Cfg.MinSpeedMps[5] := 2.5; Cfg.MaxSpeedMps[5] := 6.0;
    Cfg.MinSamples := 3;

    (* Cellule validee [1,1,1,1] puis injection hors enveloppe haute (5.0 > Max[1]=2.0) *)
    Table.Cell[1][1][1][1].Valid := TRUE;
    Table.Cell[1][1][1][1].SpeedMps := 1.5;
    Table.Cell[1][1][1][1].SampleCount := 3;
    fb(Enable := TRUE, LearnStart := TRUE, WinchId := 1, Direction := 1,
       StepNumber := 1, MeasuredSpeedMps := 5.0, MeasuredSpeedValid := TRUE,
       LoadPresent := FALSE, StableForLearn := TRUE, Config := Cfg, Table := Table);
    ASSERT_EQ(fb.CellsFilled, 0, 'Hors enveloppe haute : cellule invalidee (CellsFilled=0)');

    (* Injection sous la borne basse (0.4 < Min[1]=0.5) -> invalidation aussi *)
    Table.Cell[1][1][1][1].Valid := TRUE;
    Table.Cell[1][1][1][1].SpeedMps := 1.5;
    Table.Cell[1][1][1][1].SampleCount := 3;
    fb(Enable := TRUE, LearnStart := TRUE, WinchId := 1, Direction := 1,
       StepNumber := 1, MeasuredSpeedMps := 0.4, MeasuredSpeedValid := TRUE,
       LoadPresent := FALSE, StableForLearn := TRUE, Config := Cfg, Table := Table);
    ASSERT_EQ(fb.CellsFilled, 0, 'Sous borne basse : cellule invalidee (CellsFilled=0)');

    (* Borne exacte ==Max (2.0, inclusive) -> cellule conservee validee *)
    Table.Cell[1][1][1][1].Valid := TRUE;
    Table.Cell[1][1][1][1].SpeedMps := 1.5;
    Table.Cell[1][1][1][1].SampleCount := 3;
    fb(Enable := TRUE, LearnStart := TRUE, WinchId := 1, Direction := 1,
       StepNumber := 1, MeasuredSpeedMps := 2.0, MeasuredSpeedValid := TRUE,
       LoadPresent := FALSE, StableForLearn := TRUE, Config := Cfg, Table := Table);
    ASSERT_EQ(fb.CellsFilled, 1, 'Borne ==Max (2.0) inclusive : cellule conservee validee (1)');

    (* Borne exacte ==Min (0.5, inclusive) -> cellule conservee validee *)
    Table.Cell[1][1][1][1].Valid := TRUE;
    Table.Cell[1][1][1][1].SpeedMps := 1.5;
    Table.Cell[1][1][1][1].SampleCount := 3;
    fb(Enable := TRUE, LearnStart := TRUE, WinchId := 1, Direction := 1,
       StepNumber := 1, MeasuredSpeedMps := 0.5, MeasuredSpeedValid := TRUE,
       LoadPresent := FALSE, StableForLearn := TRUE, Config := Cfg, Table := Table);
    ASSERT_EQ(fb.CellsFilled, 1, 'Borne ==Min (0.5) inclusive : cellule conservee validee (1)');
END_TEST

TEST 'TC-T181-15e TableComplete : FALSE si une cellule manque, TRUE avec 40 cellules valides (AC6)'
VAR
    i : INT;
    j : INT;
    k : INT;
    l : INT;
END_VAR
    Cfg.MinSpeedMps[1] := 0.5; Cfg.MaxSpeedMps[1] := 2.0;
    Cfg.MinSpeedMps[2] := 1.0; Cfg.MaxSpeedMps[2] := 3.0;
    Cfg.MinSpeedMps[3] := 1.5; Cfg.MaxSpeedMps[3] := 4.0;
    Cfg.MinSpeedMps[4] := 2.0; Cfg.MaxSpeedMps[4] := 5.0;
    Cfg.MinSpeedMps[5] := 2.5; Cfg.MaxSpeedMps[5] := 6.0;
    Cfg.MinSamples := 1;

    (* Table partielle : 39 cellules valides, [2,2,2,5] manquante -> FALSE *)
    FOR i := 1 TO 2 DO
        FOR j := 1 TO 2 DO
            FOR k := 1 TO 2 DO
                FOR l := 1 TO 5 DO
                    Table.Cell[i][j][k][l].Valid := TRUE;
                END_FOR;
            END_FOR;
        END_FOR;
    END_FOR;
    Table.Cell[2][2][2][5].Valid := FALSE;

    fb(Enable := TRUE, LearnStart := FALSE, WinchId := 1, Direction := 1,
       StepNumber := 1, MeasuredSpeedMps := 1.0, MeasuredSpeedValid := TRUE,
       LoadPresent := FALSE, StableForLearn := TRUE, Config := Cfg, Table := Table);
    ASSERT_FALSE(fb.TableComplete, 'Table partielle (39/40) : TableComplete=FALSE');
    ASSERT_EQ(fb.CellsFilled, 39, 'Table partielle : CellsFilled=39');
    ASSERT_EQ(fb.CellsTotal, 40, 'CellsTotal=40 (2x2x2x5)');

    (* Table complete : 40 cellules valides -> TRUE *)
    Table.Cell[2][2][2][5].Valid := TRUE;
    fb(Enable := TRUE, LearnStart := FALSE, WinchId := 1, Direction := 1,
       StepNumber := 1, MeasuredSpeedMps := 1.0, MeasuredSpeedValid := TRUE,
       LoadPresent := FALSE, StableForLearn := TRUE, Config := Cfg, Table := Table);
    ASSERT_TRUE(fb.TableComplete, 'Table complete (40/40) : TableComplete=TRUE');
    ASSERT_EQ(fb.CellsFilled, 40, 'Table complete : CellsFilled=40');
END_TEST

TEST 'TC-T181-15f Passivite : sorties limitees au statut/diagnostic, aucune commande moteur (AC1/AC7)'
    (* La passivite (aucune sortie actionneur Relay* / Contactor* / Brake* / SpeedCmd ni
       Overspeed* / SpeedGuard* ) est verifiee par grep de l interface FB (AC1/AC7).
       Ce test confirme le comportement observable : pendant la collecte, seules les
       sorties de statut/diagnostic evoluent (Ready/Learning/LampLearn) + la Table. *)
    Cfg.MinSpeedMps[1] := 0.5; Cfg.MaxSpeedMps[1] := 2.0;
    Cfg.MinSpeedMps[2] := 1.0; Cfg.MaxSpeedMps[2] := 3.0;
    Cfg.MinSpeedMps[3] := 1.5; Cfg.MaxSpeedMps[3] := 4.0;
    Cfg.MinSpeedMps[4] := 2.0; Cfg.MaxSpeedMps[4] := 5.0;
    Cfg.MinSpeedMps[5] := 2.5; Cfg.MaxSpeedMps[5] := 6.0;
    Cfg.MinSamples := 3;

    fb(Enable := TRUE, LearnStart := TRUE, WinchId := 1, Direction := 1,
       StepNumber := 1, MeasuredSpeedMps := 1.0, MeasuredSpeedValid := TRUE,
       LoadPresent := FALSE, StableForLearn := TRUE, Config := Cfg, Table := Table);
    ASSERT_TRUE(fb.Ready, 'Enable=TRUE -> Ready=TRUE');
    ASSERT_TRUE(fb.Learning, 'Collecte active -> Learning=TRUE');
    ASSERT_TRUE(fb.LampLearn, 'Collecte active -> LampLearn=TRUE');
    ASSERT_EQ(fb.CellsTotal, 40, 'CellsTotal=40 (diagnostic)');

    (* Relache : Enable=FALSE -> Ready=FALSE, plus de collecte *)
    fb(Enable := FALSE, LearnStart := TRUE, WinchId := 1, Direction := 1,
       StepNumber := 1, MeasuredSpeedMps := 1.0, MeasuredSpeedValid := TRUE,
       LoadPresent := FALSE, StableForLearn := TRUE, Config := Cfg, Table := Table);
    ASSERT_FALSE(fb.Ready, 'Enable=FALSE -> Ready=FALSE');
    ASSERT_FALSE(fb.Learning, 'Enable=FALSE -> Learning=FALSE');
END_TEST

TEST 'TC-T181-15g Sens descente : cellule descente [1,2,1,1] ecrite, montee inchangee (AC2)'
VAR
    i : INT;
    j : INT;
    k : INT;
    l : INT;
END_VAR
    Cfg.MinSpeedMps[1] := 0.5; Cfg.MaxSpeedMps[1] := 2.0;
    Cfg.MinSpeedMps[2] := 1.0; Cfg.MaxSpeedMps[2] := 3.0;
    Cfg.MinSpeedMps[3] := 1.5; Cfg.MaxSpeedMps[3] := 4.0;
    Cfg.MinSpeedMps[4] := 2.0; Cfg.MaxSpeedMps[4] := 5.0;
    Cfg.MinSpeedMps[5] := 2.5; Cfg.MaxSpeedMps[5] := 6.0;
    Cfg.MinSamples := 1;

    (* 39 cellules valides, descente [1,2,1,1] vide. Direction=-1 -> SensIdx=2 *)
    FOR i := 1 TO 2 DO
        FOR j := 1 TO 2 DO
            FOR k := 1 TO 2 DO
                FOR l := 1 TO 5 DO
                    Table.Cell[i][j][k][l].Valid := TRUE;
                END_FOR;
            END_FOR;
        END_FOR;
    END_FOR;
    Table.Cell[1][2][1][1].Valid := FALSE;

    fb(Enable := TRUE, LearnStart := TRUE, WinchId := 1, Direction := -1,
       StepNumber := 1, MeasuredSpeedMps := 1.0, MeasuredSpeedValid := TRUE,
       LoadPresent := FALSE, StableForLearn := TRUE, Config := Cfg, Table := Table);
    ASSERT_EQ(fb.CellsFilled, 40, 'Descente : cellule descente [1,2,1,1] ecrite et validee (40)');
    ASSERT_TRUE(fb.TableComplete, 'Descente : table complete apres ecriture descente');
END_TEST

TEST 'TC-T181-15h Charge presente : cellule charge [1,1,2,1] ecrite, vide inchangee (AC2)'
VAR
    i : INT;
    j : INT;
    k : INT;
    l : INT;
END_VAR
    Cfg.MinSpeedMps[1] := 0.5; Cfg.MaxSpeedMps[1] := 2.0;
    Cfg.MinSpeedMps[2] := 1.0; Cfg.MaxSpeedMps[2] := 3.0;
    Cfg.MinSpeedMps[3] := 1.5; Cfg.MaxSpeedMps[3] := 4.0;
    Cfg.MinSpeedMps[4] := 2.0; Cfg.MaxSpeedMps[4] := 5.0;
    Cfg.MinSpeedMps[5] := 2.5; Cfg.MaxSpeedMps[5] := 6.0;
    Cfg.MinSamples := 1;

    (* 39 cellules valides, charge [1,1,2,1] vide. LoadPresent=TRUE -> ChargeIdx=2 *)
    FOR i := 1 TO 2 DO
        FOR j := 1 TO 2 DO
            FOR k := 1 TO 2 DO
                FOR l := 1 TO 5 DO
                    Table.Cell[i][j][k][l].Valid := TRUE;
                END_FOR;
            END_FOR;
        END_FOR;
    END_FOR;
    Table.Cell[1][1][2][1].Valid := FALSE;

    fb(Enable := TRUE, LearnStart := TRUE, WinchId := 1, Direction := 1,
       StepNumber := 1, MeasuredSpeedMps := 1.0, MeasuredSpeedValid := TRUE,
       LoadPresent := TRUE, StableForLearn := TRUE, Config := Cfg, Table := Table);
    ASSERT_EQ(fb.CellsFilled, 40, 'Charge : cellule charge [1,1,2,1] ecrite et validee (40)');
    ASSERT_TRUE(fb.TableComplete, 'Charge : table complete apres ecriture charge');
END_TEST

TEST 'TC-T181-15i Axe M2 (WinchId=2) : cellule [2,1,1,1] ecrite, M1 inchangee (AC2)'
VAR
    i : INT;
    j : INT;
    k : INT;
    l : INT;
END_VAR
    Cfg.MinSpeedMps[1] := 0.5; Cfg.MaxSpeedMps[1] := 2.0;
    Cfg.MinSpeedMps[2] := 1.0; Cfg.MaxSpeedMps[2] := 3.0;
    Cfg.MinSpeedMps[3] := 1.5; Cfg.MaxSpeedMps[3] := 4.0;
    Cfg.MinSpeedMps[4] := 2.0; Cfg.MaxSpeedMps[4] := 5.0;
    Cfg.MinSpeedMps[5] := 2.5; Cfg.MaxSpeedMps[5] := 6.0;
    Cfg.MinSamples := 1;

    (* 39 cellules valides, M2 [2,1,1,1] vide. WinchId=2 -> AxeIdx=2 *)
    FOR i := 1 TO 2 DO
        FOR j := 1 TO 2 DO
            FOR k := 1 TO 2 DO
                FOR l := 1 TO 5 DO
                    Table.Cell[i][j][k][l].Valid := TRUE;
                END_FOR;
            END_FOR;
        END_FOR;
    END_FOR;
    Table.Cell[2][1][1][1].Valid := FALSE;

    fb(Enable := TRUE, LearnStart := TRUE, WinchId := 2, Direction := 1,
       StepNumber := 1, MeasuredSpeedMps := 1.0, MeasuredSpeedValid := TRUE,
       LoadPresent := FALSE, StableForLearn := TRUE, Config := Cfg, Table := Table);
    ASSERT_EQ(fb.CellsFilled, 40, 'M2 : cellule [2,1,1,1] ecrite et validee (40)');
    ASSERT_TRUE(fb.TableComplete, 'M2 : table complete apres ecriture M2');
END_TEST

TEST 'TC-T181-15j Moyenne glissante + persistance RETAIN via copy-out (AC2)'
    (* Copy-out (T181-21) : apres fb(), la variable de test Table reflete les
       ecritures du FB sur la VAR_IN_OUT. On prouve ici la moyenne glissante
       (SpeedMps) et la persistance RETAIN (accumulation d'un scan a l'autre). *)
    Cfg.MinSpeedMps[1] := 0.5; Cfg.MaxSpeedMps[1] := 2.0;
    Cfg.MinSpeedMps[2] := 1.0; Cfg.MaxSpeedMps[2] := 3.0;
    Cfg.MinSpeedMps[3] := 1.5; Cfg.MaxSpeedMps[3] := 4.0;
    Cfg.MinSpeedMps[4] := 2.0; Cfg.MaxSpeedMps[4] := 5.0;
    Cfg.MinSpeedMps[5] := 2.5; Cfg.MaxSpeedMps[5] := 6.0;
    Cfg.MinSamples := 3;

    (* Cellule [1,1,1,1] vide. 1er echantillon 1.0 (plausible) -> SpeedMps=1.0, SampleCount=1 *)
    fb(Enable := TRUE, LearnStart := TRUE, WinchId := 1, Direction := 1,
       StepNumber := 1, MeasuredSpeedMps := 1.0, MeasuredSpeedValid := TRUE,
       LoadPresent := FALSE, StableForLearn := TRUE, Config := Cfg, Table := Table);
    ASSERT_EQ(Table.Cell[1][1][1][1].SampleCount, 1, '1er scan : SampleCount=1');
    ASSERT_NEAR(Table.Cell[1][1][1][1].SpeedMps, 1.0, 0.0001, '1er scan : SpeedMps=1.0');
    ASSERT_FALSE(Table.Cell[1][1][1][1].Valid, '1er scan : SampleCount<MinSamples -> Valid=FALSE');

    (* 2e echantillon 1.5 -> moyenne (1.0+1.5)/2 = 1.25, SampleCount=2 *)
    fb(Enable := TRUE, LearnStart := TRUE, WinchId := 1, Direction := 1,
       StepNumber := 1, MeasuredSpeedMps := 1.5, MeasuredSpeedValid := TRUE,
       LoadPresent := FALSE, StableForLearn := TRUE, Config := Cfg, Table := Table);
    ASSERT_EQ(Table.Cell[1][1][1][1].SampleCount, 2, '2e scan : SampleCount=2');
    ASSERT_NEAR(Table.Cell[1][1][1][1].SpeedMps, 1.25, 0.0001, '2e scan : moyenne (1.0+1.5)/2=1.25');
    ASSERT_FALSE(Table.Cell[1][1][1][1].Valid, '2e scan : SampleCount<MinSamples -> Valid=FALSE');

    (* 3e echantillon 1.5 -> moyenne (1.25*2+1.5)/3 = 1.3333, SampleCount=3 -> Valid *)
    fb(Enable := TRUE, LearnStart := TRUE, WinchId := 1, Direction := 1,
       StepNumber := 1, MeasuredSpeedMps := 1.5, MeasuredSpeedValid := TRUE,
       LoadPresent := FALSE, StableForLearn := TRUE, Config := Cfg, Table := Table);
    ASSERT_EQ(Table.Cell[1][1][1][1].SampleCount, 3, '3e scan : SampleCount=3');
    ASSERT_NEAR(Table.Cell[1][1][1][1].SpeedMps, 1.3333, 0.0001, '3e scan : moyenne (1.25*2+1.5)/3=1.3333');
    ASSERT_TRUE(Table.Cell[1][1][1][1].Valid, '3e scan : MinSamples atteint -> Valid=TRUE');
END_TEST

(* ---- test_fb_winch_symmetry.st ---- *)
(* =======================================================================
   test_fb_winch_symmetry.st -- T181-18 D11 : macro TC FB_Winch_Symmetry (F10.06)
   Observateur passif de symetrie / synchronisme M1-M2. Aucune action securite.
   Qualification : commande stable des 2 treuils, meme sens, au-dela de
   MinimumCommandTime_Ms (defaut 1000 ms) et vitesse au-dessus de MinimumSpeed_Mps.
   Les ecarts sont calcules a l arret.
   ======================================================================= *)

SETUP
VAR
    fb  : FB_Winch_Symmetry;
    Cfg : ST_fbWinch_Symmetry_Cfg;
    Dat : ST_fbWinch_Symmetry_Data;
END_VAR
END_SETUP

TEST 'TC-P10-T181-18a Cycle symetrique -> SymmetryValid et SymmetryOk'
    Cfg.MinimumCommandTime_Ms := 300;
    Cfg.MinimumSpeed_Mps := 0.05;
    Cfg.DeltaStartDelay_Ms := 100; Cfg.DeltaBrakeReleaseTime_Ms := 100;
    Cfg.DeltaBrakeApplyTime_Ms := 100; Cfg.DeltaStopDistance_Mm := 100;
    Cfg.DeltaStopTime_Ms := 200;
    fb(Reset := TRUE, M1CommandActive := FALSE, M2CommandActive := FALSE, M1Direction := 0, M2Direction := 0,
       M1BrakeCmd := FALSE, M2BrakeCmd := FALSE, M1BrakeApplied := TRUE, M2BrakeApplied := TRUE,
       M1Position_M := 0.0, M2Position_M := 0.0, M1Speed_Mps := 0.0, M2Speed_Mps := 0.0,
       SyncDeviation_M := 0.0, Config := Cfg, Data := Dat);
    fb(Reset := FALSE, M1CommandActive := TRUE, M2CommandActive := TRUE, M1Direction := 1, M2Direction := 1,
       M1BrakeCmd := TRUE, M2BrakeCmd := TRUE, M1BrakeApplied := FALSE, M2BrakeApplied := FALSE,
       M1Position_M := 0.0, M2Position_M := 0.0, M1Speed_Mps := 1.0, M2Speed_Mps := 1.0,
       SyncDeviation_M := 0.10, Config := Cfg, Data := Dat);
    ADVANCE_TIME(500000000);
    fb(Reset := FALSE, M1CommandActive := TRUE, M2CommandActive := TRUE, M1Direction := 1, M2Direction := 1,
       M1BrakeCmd := TRUE, M2BrakeCmd := TRUE, M1BrakeApplied := FALSE, M2BrakeApplied := FALSE,
       M1Position_M := 0.5, M2Position_M := 0.5, M1Speed_Mps := 1.0, M2Speed_Mps := 1.0,
       SyncDeviation_M := 0.10, Config := Cfg, Data := Dat);
    ADVANCE_TIME(500000000);
    fb(Reset := FALSE, M1CommandActive := TRUE, M2CommandActive := TRUE, M1Direction := 1, M2Direction := 1,
       M1BrakeCmd := TRUE, M2BrakeCmd := TRUE, M1BrakeApplied := FALSE, M2BrakeApplied := FALSE,
       M1Position_M := 1.0, M2Position_M := 1.0, M1Speed_Mps := 1.0, M2Speed_Mps := 1.0,
       SyncDeviation_M := 0.10, Config := Cfg, Data := Dat);
    ADVANCE_TIME(500000000);
    fb(Reset := FALSE, M1CommandActive := TRUE, M2CommandActive := TRUE, M1Direction := 1, M2Direction := 1,
       M1BrakeCmd := TRUE, M2BrakeCmd := TRUE, M1BrakeApplied := FALSE, M2BrakeApplied := FALSE,
       M1Position_M := 1.5, M2Position_M := 1.5, M1Speed_Mps := 1.0, M2Speed_Mps := 1.0,
       SyncDeviation_M := 0.10, Config := Cfg, Data := Dat);
    ADVANCE_TIME(500000000);
    fb(Reset := FALSE, M1CommandActive := FALSE, M2CommandActive := FALSE, M1Direction := 1, M2Direction := 1,
       M1BrakeCmd := FALSE, M2BrakeCmd := FALSE, M1BrakeApplied := TRUE, M2BrakeApplied := TRUE,
       M1Position_M := 2.0, M2Position_M := 2.0, M1Speed_Mps := 0.0, M2Speed_Mps := 0.0,
       SyncDeviation_M := 0.0, Config := Cfg, Data := Dat);
    ADVANCE_TIME(10000000);
    fb(Reset := FALSE, M1CommandActive := FALSE, M2CommandActive := FALSE, M1Direction := 1, M2Direction := 1,
       M1BrakeCmd := FALSE, M2BrakeCmd := FALSE, M1BrakeApplied := TRUE, M2BrakeApplied := TRUE,
       M1Position_M := 2.0, M2Position_M := 2.0, M1Speed_Mps := 0.0, M2Speed_Mps := 0.0,
       SyncDeviation_M := 0.0, Config := Cfg, Data := Dat);
    ASSERT_TRUE(fb.SymmetryValid, 'Cycle complet qualifie puis arrete -> mesure valide');
    ASSERT_TRUE(fb.SymmetryOk, 'M1 et M2 identiques -> tous les ecarts sous les seuils');
END_TEST

TEST 'TC-P10-T181-18b Reset remet les mesures a zero'
    Cfg.MinimumCommandTime_Ms := 300;
    Cfg.MinimumSpeed_Mps := 0.05;
    Cfg.DeltaStartDelay_Ms := 100; Cfg.DeltaBrakeReleaseTime_Ms := 100;
    Cfg.DeltaBrakeApplyTime_Ms := 100; Cfg.DeltaStopDistance_Mm := 100;
    Cfg.DeltaStopTime_Ms := 200;
    fb(Reset := TRUE, M1CommandActive := FALSE, M2CommandActive := FALSE, M1Direction := 0, M2Direction := 0,
       M1BrakeCmd := FALSE, M2BrakeCmd := FALSE, M1BrakeApplied := TRUE, M2BrakeApplied := TRUE,
       M1Position_M := 0.0, M2Position_M := 0.0, M1Speed_Mps := 0.0, M2Speed_Mps := 0.0,
       SyncDeviation_M := 0.0, Config := Cfg, Data := Dat);
    fb(Reset := FALSE, M1CommandActive := TRUE, M2CommandActive := TRUE, M1Direction := 1, M2Direction := 1,
       M1BrakeCmd := TRUE, M2BrakeCmd := TRUE, M1BrakeApplied := FALSE, M2BrakeApplied := FALSE,
       M1Position_M := 0.0, M2Position_M := 0.0, M1Speed_Mps := 1.0, M2Speed_Mps := 1.0,
       SyncDeviation_M := 0.40, Config := Cfg, Data := Dat);
    ADVANCE_TIME(600000000);
    fb(Reset := FALSE, M1CommandActive := TRUE, M2CommandActive := TRUE, M1Direction := 1, M2Direction := 1,
       M1BrakeCmd := TRUE, M2BrakeCmd := TRUE, M1BrakeApplied := FALSE, M2BrakeApplied := FALSE,
       M1Position_M := 0.6, M2Position_M := 0.6, M1Speed_Mps := 1.0, M2Speed_Mps := 1.0,
       SyncDeviation_M := 0.40, Config := Cfg, Data := Dat);
    ADVANCE_TIME(600000000);
    fb(Reset := FALSE, M1CommandActive := TRUE, M2CommandActive := TRUE, M1Direction := 1, M2Direction := 1,
       M1BrakeCmd := TRUE, M2BrakeCmd := TRUE, M1BrakeApplied := FALSE, M2BrakeApplied := FALSE,
       M1Position_M := 1.2, M2Position_M := 1.2, M1Speed_Mps := 1.0, M2Speed_Mps := 1.0,
       SyncDeviation_M := 0.40, Config := Cfg, Data := Dat);
    fb(Reset := TRUE, M1CommandActive := FALSE, M2CommandActive := FALSE, M1Direction := 0, M2Direction := 0,
       M1BrakeCmd := FALSE, M2BrakeCmd := FALSE, M1BrakeApplied := TRUE, M2BrakeApplied := TRUE,
       M1Position_M := 0.0, M2Position_M := 0.0, M1Speed_Mps := 0.0, M2Speed_Mps := 0.0,
       SyncDeviation_M := 0.0, Config := Cfg, Data := Dat);
    ASSERT_EQ(Dat.DeltaStartDelay_Ms, 0, 'Reset -> DeltaStartDelay_Ms remis a 0');
    ASSERT_FALSE(Dat.MaxSyncDeviation_M > 0.0, 'Reset -> MaxSyncDeviation_M remis a 0');
END_TEST

TEST 'TC-P10-T181-18c Non qualifie si un seul treuil commande'
    Cfg.MinimumCommandTime_Ms := 300;
    Cfg.MinimumSpeed_Mps := 0.05;
    Cfg.DeltaStartDelay_Ms := 100; Cfg.DeltaBrakeReleaseTime_Ms := 100;
    Cfg.DeltaBrakeApplyTime_Ms := 100; Cfg.DeltaStopDistance_Mm := 100;
    Cfg.DeltaStopTime_Ms := 200;
    fb(Reset := TRUE, M1CommandActive := FALSE, M2CommandActive := FALSE, M1Direction := 0, M2Direction := 0,
       M1BrakeCmd := FALSE, M2BrakeCmd := FALSE, M1BrakeApplied := TRUE, M2BrakeApplied := TRUE,
       M1Position_M := 0.0, M2Position_M := 0.0, M1Speed_Mps := 0.0, M2Speed_Mps := 0.0,
       SyncDeviation_M := 0.0, Config := Cfg, Data := Dat);
    fb(Reset := FALSE, M1CommandActive := TRUE, M2CommandActive := FALSE, M1Direction := 1, M2Direction := 0,
       M1BrakeCmd := TRUE, M2BrakeCmd := FALSE, M1BrakeApplied := FALSE, M2BrakeApplied := TRUE,
       M1Position_M := 0.0, M2Position_M := 0.0, M1Speed_Mps := 1.0, M2Speed_Mps := 0.0,
       SyncDeviation_M := 0.30, Config := Cfg, Data := Dat);
    ADVANCE_TIME(1500000000);
    fb(Reset := FALSE, M1CommandActive := TRUE, M2CommandActive := FALSE, M1Direction := 1, M2Direction := 0,
       M1BrakeCmd := TRUE, M2BrakeCmd := FALSE, M1BrakeApplied := FALSE, M2BrakeApplied := TRUE,
       M1Position_M := 1.5, M2Position_M := 0.0, M1Speed_Mps := 1.0, M2Speed_Mps := 0.0,
       SyncDeviation_M := 0.30, Config := Cfg, Data := Dat);
    ASSERT_FALSE(fb.SymmetryValid, 'Un seul treuil commande -> jamais qualifie');
END_TEST

(* ---- test_fb_winchdirectioninterlock.st ---- *)
(* =======================================================================
   test_fb_winchdirectioninterlock.st — T181-18 D11 : macro TC FB_WinchDirectionInterlock
   ======================================================================= *)

SETUP
VAR
    fb : FB_WinchDirectionInterlock;
END_VAR
END_SETUP

TEST 'TC-P10-T181-18a Premier sens depuis le neutre : adoption immediate'
    fb(Enable := TRUE, EnableRising := FALSE, Reset := FALSE, ReqDirection := 1, ChangeDelayUp := T#900ms, ChangeDelayDown := T#400ms);
    ASSERT_EQ(fb.CommandedDirection, 1, 'Adoption immediate du premier sens');
    ASSERT_FALSE(fb.DirectionChangePending, 'Pas de pending');
END_TEST

TEST 'TC-P10-T181-18b Reprise du meme sens apres neutre : immediate'
    fb(Enable := TRUE, EnableRising := FALSE, Reset := FALSE, ReqDirection := 1, ChangeDelayUp := T#900ms, ChangeDelayDown := T#400ms);
    fb(Enable := TRUE, EnableRising := FALSE, Reset := FALSE, ReqDirection := 0, ChangeDelayUp := T#900ms, ChangeDelayDown := T#400ms);
    ASSERT_EQ(fb.CommandedDirection, 0, 'Retour au neutre');
    fb(Enable := TRUE, EnableRising := FALSE, Reset := FALSE, ReqDirection := 1, ChangeDelayUp := T#900ms, ChangeDelayDown := T#400ms);
    ASSERT_EQ(fb.CommandedDirection, 1, 'Reprise du meme sens : immediate');
    ASSERT_FALSE(fb.DirectionChangePending, 'Pas de pending');
END_TEST

TEST 'TC-P10-T181-18c Reprise du sens oppose : adoption seulement apres le delai'
    fb(Enable := TRUE, EnableRising := FALSE, Reset := FALSE, ReqDirection := 1, ChangeDelayUp := T#900ms, ChangeDelayDown := T#400ms);
    fb(Enable := TRUE, EnableRising := FALSE, Reset := FALSE, ReqDirection := 0, ChangeDelayUp := T#900ms, ChangeDelayDown := T#400ms);
    fb(Enable := TRUE, EnableRising := FALSE, Reset := FALSE, ReqDirection := -1, ChangeDelayUp := T#900ms, ChangeDelayDown := T#400ms);
    ASSERT_EQ(fb.CommandedDirection, 0, 'Pas encore adopte (pending)');
    ASSERT_TRUE(fb.DirectionChangePending, 'Pending actif avant le delai');
    ADVANCE_TIME(400000000);
    fb(Enable := TRUE, EnableRising := FALSE, Reset := FALSE, ReqDirection := -1, ChangeDelayUp := T#900ms, ChangeDelayDown := T#400ms);
    ASSERT_EQ(fb.CommandedDirection, -1, 'Sens oppose adopte apres ChangeDelayDown');
    ASSERT_FALSE(fb.DirectionChangePending, 'Pending termine');
END_TEST

TEST 'TC-P10-T181-18d ReqDirection=0 force le neutre'
    fb(Enable := TRUE, EnableRising := FALSE, Reset := FALSE, ReqDirection := 1, ChangeDelayUp := T#900ms, ChangeDelayDown := T#400ms);
    fb(Enable := TRUE, EnableRising := FALSE, Reset := FALSE, ReqDirection := 0, ChangeDelayUp := T#900ms, ChangeDelayDown := T#400ms);
    ASSERT_EQ(fb.CommandedDirection, 0, 'Neutre commande');
    ASSERT_FALSE(fb.DirectionChangePending, 'Pas de pending au neutre');
END_TEST

(* ---- test_fb_winchloadestimator.st ---- *)
(* =======================================================================
   test_fb_winchloadestimator.st — T181-18 D11 : macro TC FB_WinchLoadEstimator
   Estimateur informatif (aucune action securite). Couvre : gate, classement
   de vitesse par bande + hysteresis, direction montee/descente, validation table.
   (La lecture de la matrice 5x5 elle-meme n'est pas asserted ici : passthrough,
   et le harnais STruCpp ne supporte pas l'indexation [i][j] d'un ARRAY OF ARRAY.)
   ======================================================================= *)

SETUP
VAR
    fb  : FB_WinchLoadEstimator;
    Spd : ST_fbWinchLoadEstimator_SpeedCfg;
    Tbl : ST_fbWinchLoadEstimator_Table;
END_VAR
END_SETUP

TEST 'TC-P10-T181-18a Gate : Enable FALSE -> sorties neutres'
    Spd.MaxMeasuredSpeedMps := 2.0;
    Spd.SpeedBandMaxMps[1] := 0.4; Spd.SpeedBandMaxMps[2] := 0.8; Spd.SpeedBandMaxMps[3] := 1.2;
    Spd.SpeedBandMaxMps[4] := 1.6; Spd.SpeedBandMaxMps[5] := 2.0;
    Spd.SpeedBandHysteresisMps := 0.05;
    fb(Enable := FALSE, PowerContactorEngaged := TRUE, ActiveSpeedStep := 3,
       MeasuredSpeedMps := 0.5, MeasuredSpeedSignedMps := 0.5,
       SpeedConfig := Spd, LoadTable := Tbl);
    ASSERT_FALSE(fb.Ready, 'Enable FALSE -> Ready FALSE');
    ASSERT_EQ(fb.SpeedBand, 0, 'Enable FALSE -> SpeedBand 0');
    ASSERT_EQ(fb.EstimatedLoadPct, 0.0, 'Enable FALSE -> estimation 0');
END_TEST

TEST 'TC-P10-T181-18b Classement vitesse : 0.5 m/s -> bande 2, montee'
    Spd.MaxMeasuredSpeedMps := 2.0;
    Spd.SpeedBandMaxMps[1] := 0.4; Spd.SpeedBandMaxMps[2] := 0.8; Spd.SpeedBandMaxMps[3] := 1.2;
    Spd.SpeedBandMaxMps[4] := 1.6; Spd.SpeedBandMaxMps[5] := 2.0;
    Spd.SpeedBandHysteresisMps := 0.05;
    Tbl.IsConfigured := TRUE;
    fb(Enable := TRUE, PowerContactorEngaged := TRUE, ActiveSpeedStep := 2,
       MeasuredSpeedMps := 0.5, MeasuredSpeedSignedMps := 0.5,
       SpeedConfig := Spd, LoadTable := Tbl);
    ASSERT_EQ(fb.SpeedBand, 2, 'Vitesse 0.5 m/s (entre 0.4 et 0.8) -> bande 2');
    ASSERT_TRUE(fb.Ascending, 'Vitesse signee positive -> montee');
    ASSERT_TRUE(fb.Configured, 'Table validee -> Configured TRUE');
    ASSERT_TRUE(fb.Ready, 'Nominal -> Ready TRUE');
END_TEST

TEST 'TC-P10-T181-18c Classement vitesse : 1.5 m/s -> bande 4'
    Spd.MaxMeasuredSpeedMps := 2.0;
    Spd.SpeedBandMaxMps[1] := 0.4; Spd.SpeedBandMaxMps[2] := 0.8; Spd.SpeedBandMaxMps[3] := 1.2;
    Spd.SpeedBandMaxMps[4] := 1.6; Spd.SpeedBandMaxMps[5] := 2.0;
    Spd.SpeedBandHysteresisMps := 0.05;
    fb(Enable := TRUE, PowerContactorEngaged := TRUE, ActiveSpeedStep := 4,
       MeasuredSpeedMps := 1.5, MeasuredSpeedSignedMps := 1.5,
       SpeedConfig := Spd, LoadTable := Tbl);
    ASSERT_EQ(fb.SpeedBand, 4, 'Vitesse 1.5 m/s (entre 1.2 et 1.6) -> bande 4');
END_TEST

TEST 'TC-P10-T181-18d Descente : aucune estimation de charge'
    Spd.MaxMeasuredSpeedMps := 2.0;
    Spd.SpeedBandMaxMps[1] := 0.4; Spd.SpeedBandMaxMps[2] := 0.8; Spd.SpeedBandMaxMps[3] := 1.2;
    Spd.SpeedBandMaxMps[4] := 1.6; Spd.SpeedBandMaxMps[5] := 2.0;
    Spd.SpeedBandHysteresisMps := 0.05;
    Tbl.IsConfigured := TRUE;
    fb(Enable := TRUE, PowerContactorEngaged := TRUE, ActiveSpeedStep := 2,
       MeasuredSpeedMps := 0.5, MeasuredSpeedSignedMps := -0.5,
       SpeedConfig := Spd, LoadTable := Tbl);
    ASSERT_FALSE(fb.Ascending, 'Vitesse signee negative -> descente');
    ASSERT_EQ(fb.EstimatedLoadPct, 0.0, 'Descente : estimation non produite');
END_TEST

TEST 'TC-P10-T181-18e Vitesse mesuree negative -> defaut latche, bande 0'
    Spd.MaxMeasuredSpeedMps := 2.0;
    Spd.SpeedBandMaxMps[1] := 0.4; Spd.SpeedBandMaxMps[2] := 0.8; Spd.SpeedBandMaxMps[3] := 1.2;
    Spd.SpeedBandMaxMps[4] := 1.6; Spd.SpeedBandMaxMps[5] := 2.0;
    Spd.SpeedBandHysteresisMps := 0.05;
    fb(Enable := TRUE, PowerContactorEngaged := TRUE, ActiveSpeedStep := 2,
       MeasuredSpeedMps := -0.1, MeasuredSpeedSignedMps := -0.1,
       SpeedConfig := Spd, LoadTable := Tbl);
    ASSERT_EQ(fb.SpeedBand, 0, 'Vitesse mesuree < 0 -> bande 0');
    (* Le socle latche la cause au scan suivant (Active pose apres l'appel FB_FaultCore). *)
    fb(Enable := TRUE, PowerContactorEngaged := TRUE, ActiveSpeedStep := 2,
       MeasuredSpeedMps := -0.1, MeasuredSpeedSignedMps := -0.1,
       SpeedConfig := Spd, LoadTable := Tbl);
    ASSERT_TRUE(fb.Fault.Latched, 'Vitesse mesuree < 0 -> defaut latche');
END_TEST
